Fanuc KAREL source: kc00015.KL

-- PROVISIONAL review KL for V1013-1; original PC SHA256 75d767cec6c0b88762bc50b26254a4bff148af2eaa150918908cc336ec29db4d
-- Incomplete behavior may be omitted. Consult companion uncertainty JSON. Do not deploy.
PROGRAM KC00015
%NOLOCKGROUP
BEGIN
  -- UNRESOLVED_PC offsets 5-12; opcodes 9D,23
  -- UNRESOLVED_PC offsets 17-47; opcodes 27,22,22,27,9D,31,7E,4A
  -- UNRESOLVED_PC offsets 52-56; opcodes 7F
END KC00015
